FUNCTION_BLOCK BATCH_FILLING (* Solvability control: ecc_persistent form, designed by hand. Never shown to a model. *)
  (* Standard: 61499-2 *)
  (* Version 1.0, 2026-11-06, st2fb *)
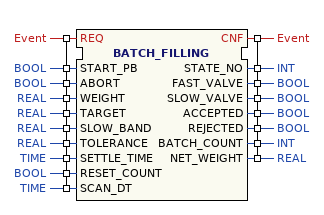
  EVENT_INPUT
    REQ WITH START_PB, ABORT, WEIGHT, TARGET, SLOW_BAND, TOLERANCE, SETTLE_TIME, RESET_COUNT, SCAN_DT;
  END_EVENT
  EVENT_OUTPUT
    CNF WITH STATE_NO, FAST_VALVE, SLOW_VALVE, ACCEPTED, REJECTED, BATCH_COUNT, NET_WEIGHT;
  END_EVENT
  VAR_INPUT
    START_PB : BOOL;
    ABORT : BOOL;
    WEIGHT : REAL;
    TARGET : REAL;
    SLOW_BAND : REAL;
    TOLERANCE : REAL;
    SETTLE_TIME : TIME;
    RESET_COUNT : BOOL;
    SCAN_DT : TIME;
  END_VAR
  VAR_OUTPUT
    STATE_NO : INT;
    FAST_VALVE : BOOL;
    SLOW_VALVE : BOOL;
    ACCEPTED : BOOL;
    REJECTED : BOOL;
    BATCH_COUNT : INT;
    NET_WEIGHT : REAL;
  END_VAR
  VAR
    TARE : REAL;
    COUNT_PULSE : BOOL;
    ST2FB_NOW : TIME;
    SETTLE_TIMER_IN : BOOL;
    SETTLE_TIMER_PT : TIME;
    SETTLE_TIMER_Q : BOOL;
    SETTLE_TIMER_ET : TIME;
    SETTLE_TIMER_STATE : INT;
    SETTLE_TIMER_PREV_IN : BOOL;
    SETTLE_TIMER_START_TIME : TIME;
    COUNTER_CU : BOOL;
    COUNTER_R : BOOL;
    COUNTER_PV : INT;
    COUNTER_Q : BOOL;
    COUNTER_CV : INT;
    COUNTER_CU_T_Q : BOOL;
    COUNTER_CU_T_M : BOOL;
    START_EDGE_CLK : BOOL;
    START_EDGE_Q : BOOL;
    START_EDGE_M : BOOL;
  END_VAR
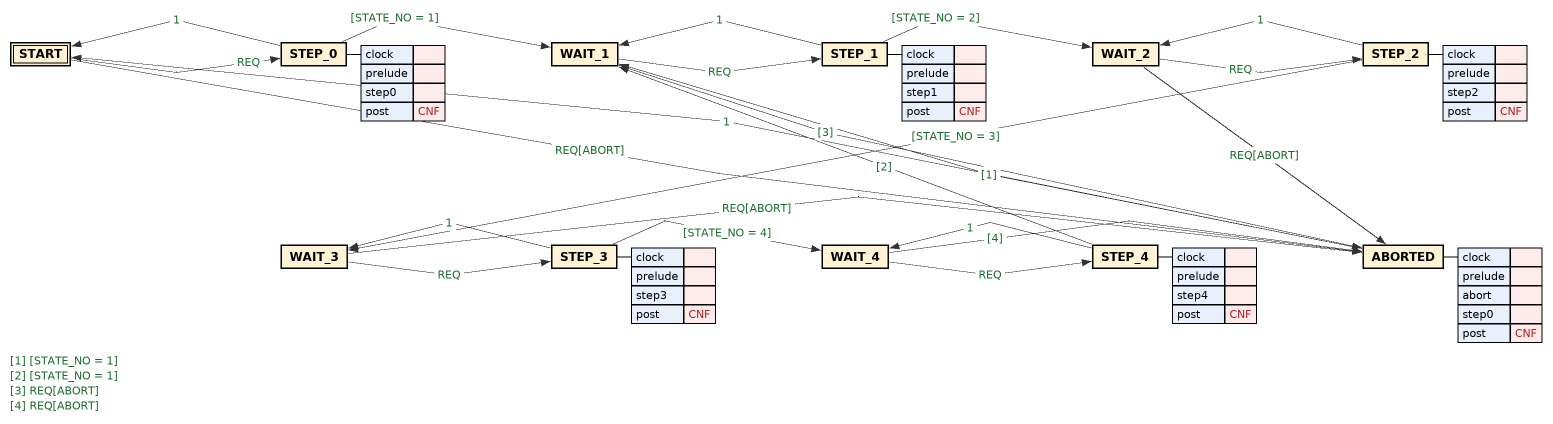
  EC_STATES
    START;
    STEP_0 : clock, prelude, step0, post -> CNF;
    WAIT_1;
    STEP_1 : clock, prelude, step1, post -> CNF;
    WAIT_2;
    STEP_2 : clock, prelude, step2, post -> CNF;
    WAIT_3;
    STEP_3 : clock, prelude, step3, post -> CNF;
    WAIT_4;
    STEP_4 : clock, prelude, step4, post -> CNF;
    ABORTED : clock, prelude, abort, step0, post -> CNF;
  END_STATES
  EC_TRANSITIONS
    START TO ABORTED := REQ[ABORT];
    START TO STEP_0 := REQ;
    WAIT_1 TO ABORTED := REQ[ABORT];
    WAIT_1 TO STEP_1 := REQ;
    WAIT_2 TO ABORTED := REQ[ABORT];
    WAIT_2 TO STEP_2 := REQ;
    WAIT_3 TO ABORTED := REQ[ABORT];
    WAIT_3 TO STEP_3 := REQ;
    WAIT_4 TO ABORTED := REQ[ABORT];
    WAIT_4 TO STEP_4 := REQ;
    STEP_0 TO WAIT_1 := [STATE_NO = 1];
    STEP_0 TO START := 1;
    ABORTED TO WAIT_1 := [STATE_NO = 1];
    ABORTED TO START := 1;
    STEP_1 TO WAIT_2 := [STATE_NO = 2];
    STEP_1 TO WAIT_1 := 1;
    STEP_2 TO WAIT_3 := [STATE_NO = 3];
    STEP_2 TO WAIT_2 := 1;
    STEP_3 TO WAIT_4 := [STATE_NO = 4];
    STEP_3 TO WAIT_3 := 1;
    STEP_4 TO WAIT_1 := [STATE_NO = 1];
    STEP_4 TO WAIT_4 := 1;
  END_TRANSITIONS
  ALGORITHM clock IN ST:
ST2FB_NOW := ST2FB_NOW + SCAN_DT;
  END_ALGORITHM
  ALGORITHM prelude IN ST:
START_EDGE_CLK := START_PB;
START_EDGE_Q := START_EDGE_CLK AND NOT START_EDGE_M;
START_EDGE_M := START_EDGE_CLK;
NET_WEIGHT := WEIGHT - TARE;
FAST_VALVE := FALSE;
SLOW_VALVE := FALSE;
COUNT_PULSE := FALSE;
  END_ALGORITHM
  ALGORITHM abort IN ST:
STATE_NO := 0;
ACCEPTED := FALSE;
REJECTED := FALSE;
  END_ALGORITHM
  ALGORITHM step0 IN ST:
IF START_EDGE_Q AND NOT ABORT THEN
  TARE := WEIGHT;
  NET_WEIGHT := 0.0;
  ACCEPTED := FALSE;
  REJECTED := FALSE;
  STATE_NO := 1;
END_IF;
  END_ALGORITHM
  ALGORITHM step1 IN ST:
FAST_VALVE := TRUE;
SLOW_VALVE := TRUE;
IF NET_WEIGHT >= TARGET - SLOW_BAND THEN
  STATE_NO := 2;
END_IF;
  END_ALGORITHM
  ALGORITHM step2 IN ST:
SLOW_VALVE := TRUE;
IF NET_WEIGHT >= TARGET THEN
  STATE_NO := 3;
END_IF;
  END_ALGORITHM
  ALGORITHM step3 IN ST:
IF SETTLE_TIMER_Q THEN
  IF NET_WEIGHT >= TARGET - TOLERANCE AND NET_WEIGHT <= TARGET + TOLERANCE THEN
    ACCEPTED := TRUE;
    COUNT_PULSE := TRUE;
  ELSE
    REJECTED := TRUE;
  END_IF;
  STATE_NO := 4;
END_IF;
  END_ALGORITHM
  ALGORITHM step4 IN ST:
IF START_EDGE_Q THEN
  TARE := WEIGHT;
  NET_WEIGHT := 0.0;
  ACCEPTED := FALSE;
  REJECTED := FALSE;
  STATE_NO := 1;
END_IF;
  END_ALGORITHM
  ALGORITHM post IN ST:
SETTLE_TIMER_IN := STATE_NO = 3;
SETTLE_TIMER_PT := SETTLE_TIME;
IF SETTLE_TIMER_STATE = 0 AND NOT SETTLE_TIMER_PREV_IN AND SETTLE_TIMER_IN THEN
  SETTLE_TIMER_STATE := 1;
  SETTLE_TIMER_Q := FALSE;
  SETTLE_TIMER_START_TIME := ST2FB_NOW;
ELSE
  IF NOT SETTLE_TIMER_IN THEN
    SETTLE_TIMER_ET := T#0s;
    SETTLE_TIMER_Q := FALSE;
    SETTLE_TIMER_STATE := 0;
  ELSIF SETTLE_TIMER_STATE = 1 THEN
    IF SETTLE_TIMER_START_TIME + SETTLE_TIMER_PT <= ST2FB_NOW THEN
      SETTLE_TIMER_STATE := 2;
      SETTLE_TIMER_Q := TRUE;
      SETTLE_TIMER_ET := SETTLE_TIMER_PT;
    ELSE
      SETTLE_TIMER_ET := ST2FB_NOW - SETTLE_TIMER_START_TIME;
    END_IF;
  END_IF;
END_IF;
SETTLE_TIMER_PREV_IN := SETTLE_TIMER_IN;
COUNTER_CU := COUNT_PULSE;
COUNTER_R := RESET_COUNT;
COUNTER_PV := 1000;
COUNTER_CU_T_Q := COUNTER_CU AND NOT COUNTER_CU_T_M;
COUNTER_CU_T_M := COUNTER_CU;
IF COUNTER_R THEN
  COUNTER_CV := 0;
ELSIF COUNTER_CU_T_Q AND COUNTER_CV < COUNTER_PV THEN
  COUNTER_CV := COUNTER_CV + 1;
END_IF;
COUNTER_Q := COUNTER_CV >= COUNTER_PV;
BATCH_COUNT := COUNTER_CV;
  END_ALGORITHM
END_FUNCTION_BLOCK
